// Motion model of one mocked axis (telescope state machine mock rig, BROTLib plan 2026-10-21-telescope-state-machine-unification).
// One call = one PLC scan of the axis part. Enable -> Ready after nReadyScans, homing -> calibrated after nHomeScans, a rising
// bMove -> InMotion for nMoveScans, then MoveDone for one scan and the position is the target. Only the levels the telescope
// writes are inputs; nothing here touches an MC_* block. Same model as MONETcommonTests.
FUNCTION_BLOCK FB_AxisMockCore
VAR_INPUT
	bEnable			: BOOL;
	bHome			: BOOL;
	bMove			: BOOL;
	bStop			: BOOL;		// the StopAxis level: a rising edge is a stop request (MC_Stop)
	fTarget			: LREAL;
	nReadyScans		: UINT := 2;
	nHomeScans		: UINT := 3;
	nMoveScans		: UINT := 4;
	nStopScans		: UINT := 3;
	bSuppressStopDone	: BOOL;	// the stop ends at rest but bStopDone is never reported (a lost Done, #120)
	nStartScans		: UINT;		// scans between the move command and the axis reporting InMotion (the NC takes a few cycles; 0 = at once). #92
END_VAR
VAR_OUTPUT
	bReady			: BOOL;
	bCalibrated		: BOOL;
	bHoming			: BOOL;
	bInMotion		: BOOL;
	bStandStill		: BOOL := TRUE;
	bMoveDone		: BOOL;		// one scan
	bStopping		: BOOL;
	bStopDone		: BOOL;		// one scan
	nStopEdges		: UINT;		// rising edges of bStop, i.e. MC_Stop requests
	fPosition		: LREAL;
END_VAR
VAR
	nReadyCount		: UINT;
	nHomeCount		: UINT;
	nMoveCount		: UINT;
	nStopCount		: UINT;
	nStartCount		: UINT;
	bStartPending	: BOOL;
	rtMove			: R_TRIG;
	rtStop			: R_TRIG;
END_VAR

bMoveDone := FALSE;
bStopDone := FALSE;

// a stop request aborts a running move where it is (the model has no interpolation: the position stays) and takes
// nStopScans scans, then reports Done for one scan
rtStop(CLK := bStop);
IF rtStop.Q THEN
	nStopEdges := nStopEdges + 1;
	bStopping := TRUE;
	nStopCount := 0;
	bInMotion := FALSE;
	bStartPending := FALSE;
END_IF
IF bStopping THEN
	nStopCount := nStopCount + 1;
	IF nStopCount >= nStopScans THEN
		bStopping := FALSE;
		bStopDone := NOT bSuppressStopDone;
	END_IF
END_IF

IF bEnable THEN
	IF nReadyCount >= nReadyScans THEN
		bReady := TRUE;
	ELSE
		nReadyCount := nReadyCount + 1;
	END_IF
ELSE
	nReadyCount := 0;
	bReady := FALSE;
END_IF

IF bHome AND bReady AND NOT bCalibrated THEN
	bHoming := TRUE;
	nHomeCount := nHomeCount + 1;
	IF nHomeCount >= nHomeScans THEN
		bCalibrated := TRUE;
		bHoming := FALSE;
		nHomeCount := 0;
	END_IF
ELSE
	bHoming := FALSE;
END_IF

rtMove(CLK := bMove);
IF rtMove.Q AND bReady AND bCalibrated AND NOT bStopping THEN
	IF nStartScans = 0 THEN
		bInMotion := TRUE;
		nMoveCount := 0;
	ELSE
		// the move command is out, the axis still reports StandStill until the NC has started it (#92)
		bStartPending := TRUE;
		nStartCount := 0;
	END_IF
ELSIF bStartPending THEN
	nStartCount := nStartCount + 1;
	IF nStartCount >= nStartScans THEN
		bStartPending := FALSE;
		bInMotion := TRUE;
		nMoveCount := 0;
	END_IF
END_IF
IF bInMotion THEN
	nMoveCount := nMoveCount + 1;
	IF nMoveCount >= nMoveScans THEN
		fPosition := fTarget;
		bInMotion := FALSE;
		bMoveDone := TRUE;
	END_IF
END_IF

bStandStill := NOT bInMotion AND NOT bHoming AND NOT bStopping;

END_FUNCTION_BLOCK

(* stored: Version 1.1.0.1, ProductVersion 3.1.4024.15
   POU FB_AxisMockCore: Id {f878c1e1-168b-48b7-98af-f8744b9b9559}, SpecialFunc None *)
